(* IEC 61131-3 sources: SRCI_CLIENT_PLC/RobotLibrary/Library/POUs/General/MC_UserLogin/Structures, 4 files *)

(* ---- UserLoginOutCmd.st ---- *)
{attribute 'pack_mode' := '1'}
// -------------------------------------------------------------------------
//  SRCI Robot Library
// -------------------------------------------------------------------------
//
//  Object:      UserLoginOutCmd
//  Author:      Thorsten Brach
//  Date:        2024-06-30
//
//  Description:
//
//
//  Copyright:
//    (C) 2024 Thorsten Brach. All rights reserved
//             Licensed under the MIT License.
//
//  Disclaimer:
//    This project is provided without any guarantee and can be used for
//    private and commercial purposes. Any use is at the user’s
//    own risk and responsibility.
//
// -------------------------------------------------------------------------
TYPE UserLoginOutCmd :
STRUCT
END_STRUCT
END_TYPE

(* ---- UserLoginParCmd.st ---- *)
{attribute 'pack_mode' := '1'}
// -------------------------------------------------------------------------
//  SRCI Robot Library
// -------------------------------------------------------------------------
//
//  Object:      UserLoginParCmd
//  Author:      Thorsten Brach
//  Date:        2024-06-30
//
//  Description:
//
//
//  Copyright:
//    (C) 2024 Thorsten Brach. All rights reserved
//             Licensed under the MIT License.
//
//  Disclaimer:
//    This project is provided without any guarantee and can be used for
//    private and commercial purposes. Any use is at the user’s
//    own risk and responsibility.
//
// -------------------------------------------------------------------------
TYPE UserLoginParCmd :
STRUCT
  /// Defines the logon type (at least one option must be supported)
  Mode            : LogonMode;
  /// Defines the user password.
  Password        : STRING(50);
  /// Defines the name of the operator
  Username        : STRING(50);
  /// Defines the level ID of the operator (default: 0)
  LevelID         : SINT;
END_STRUCT
END_TYPE

(* ---- UserLoginRecvData.st ---- *)
{attribute 'pack_mode' := '1'}
// -------------------------------------------------------------------------
//  SRCI Robot Library
// -------------------------------------------------------------------------
//
//  Object:      UserLoginRecvData
//  Author:      Thorsten Brach
//  Date:        2024-06-30
//
//  Description:
//
//
//  Copyright:
//    (C) 2024 Thorsten Brach. All rights reserved
//             Licensed under the MIT License.
//
//  Disclaimer:
//    This project is provided without any guarantee and can be used for
//    private and commercial purposes. Any use is at the user’s
//    own risk and responsibility.
//
// -------------------------------------------------------------------------
TYPE UserLoginRecvData EXTENDS RspHeader :
STRUCT
END_STRUCT
END_TYPE

(* ---- UserLoginSendData.st ---- *)
{attribute 'pack_mode' := '1'}
// -------------------------------------------------------------------------
//  SRCI Robot Library
// -------------------------------------------------------------------------
//
//  Object:      UserLoginSendData
//  Author:      Thorsten Brach
//  Date:        2024-06-30
//
//  Description:
//
//
//  Copyright:
//    (C) 2024 Thorsten Brach. All rights reserved
//             Licensed under the MIT License.
//
//  Disclaimer:
//    This project is provided without any guarantee and can be used for
//    private and commercial purposes. Any use is at the user’s
//    own risk and responsibility.
//
// -------------------------------------------------------------------------
TYPE UserLoginSendData EXTENDS CmdHeader:
STRUCT
  /// Defines the logon type (at least one option must be supported)
  Mode            : LogonMode;
  /// Defines the level ID of the operator (default: 0)
  LevelID         : SINT;
  /// Defines the user password.
  Password        : STRING(50);
  /// Defines the name of the operator
  Username        : STRING(50);
END_STRUCT
END_TYPE
